DATA_BLOCK "iKraanSim1"
{ S7_Optimized_Access := 'TRUE' }
VERSION : 0.1
NON_RETAIN
"FB_KraanSim"

BEGIN

END_DATA_BLOCK

DATA_BLOCK "iMes"
{ S7_Optimized_Access := 'TRUE' }
VERSION : 0.1
NON_RETAIN
"FB_Mes"

BEGIN

END_DATA_BLOCK

DATA_BLOCK "iKraanSim2"
{ S7_Optimized_Access := 'TRUE' }
VERSION : 0.1
NON_RETAIN
"FB_KraanSim"

BEGIN

END_DATA_BLOCK

